Staubli VAL3: refreshList.pgx

program refreshList()
  local num l_i
begin
  for l_i = 0 to size(sFrameList)-1
    sFrameList[l_i]=toString("",l_i)+","+savedata:fFrameItem[l_i].sName
  endFor

  for l_i = 0 to size(sToolList)-1
    sToolList[l_i]=toString("",l_i)+","+savedata:tToolItem[l_i].sName
  endFor
end
